Fanuc KAREL source: KT00547.KL

PROGRAM KT00547
%NOLOCKGROUP
VAR
  P1: JOINTPOS
  P2: XYZWPREXT
  OUT: JOINTPOS
BEGIN
    P2.Y = 2.0
  OUT = P1 : P2
END KT00547
